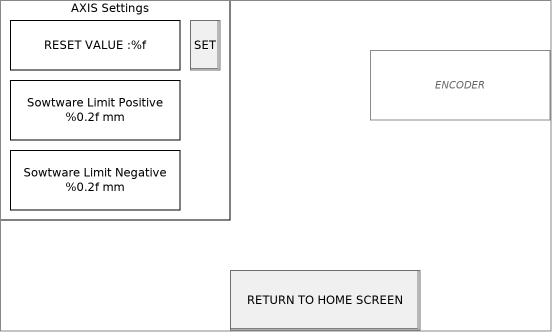
VISUALIZATION AXIS  // 552x332
    Rectangle (-10,0 240x220), "AXIS Settings"
    Rectangle (10,20 170x50), "RESET VALUE :%f", text variable: MAIN.Track.PositionResetValue
        OnMouseDown: write the text variable via VisuDialogs.Numpad, title 'Reset Value'
    Button (190,20 30x50), "SET"
        tap MAIN.Track.PositionReset
    Rectangle (10,80 170x60), "Sowtware Limit Positive %0.2f mm", text variable: MAIN.Track.LimitPos
    Rectangle (10,150 170x60), "Sowtware Limit Negative %0.2f mm", text variable: MAIN.Track.LimitNeg
    Button (230,270 190x60), "RETURN TO HOME SCREEN"
        OnMouseUp: change screen: TC_VISU
    Frame (370,50 180x70)
        shows ENCODER()
END_VISUALIZATION

(* stored: Version 1.1.0.1, ProductVersion 3.1.4024.16
   Visu AXIS: Id {baee7f2a-0daa-46cf-b43d-8143d2e5619c} *)
